Fanuc KAREL source: ka00027.KL

PROGRAM KA00027
%STACKSIZE=65535
%PRIORITY=65535
%NOLOCKGROUP
VAR
SRC : BOOLEAN
DST : BOOLEAN
BEGIN
SRC=TRUE
DST=SRC
END KA00027
